(* IEC 61131-3 sources: Caravan/Archiv/12-04-19/Stations/MachineControl/MachineControl/Class/SafetyCDIAS_Base (part 6) *)

END_FUNCTION

FUNCTION VIRTUAL SafetyCDIAS_Base::GetChannelInfo
	VAR_INPUT
		pErrorMemUser 	: ^UINT;
		pErrorMem 	: ^USINT;
		ErrorDataLength 	: INT;
	END_VAR
	VAR_OUTPUT
		StateReady 	: BOOL;
	END_VAR
  VAR
  	i   : INT;
  END_VAR

  StateReady := DiagVars.UserErrorInfoReady;

  if StateReady then
    //copy error values in UserArray
    for i := 0 to ErrorDataLength-1 do

      pErrorMemUser^ := pErrorMem^;

      //set pointer to next entry
      pErrorMemUser += sizeof(UINT);
      pErrorMem += sizeof(USINT);
    end_for;
  end_if;

END_FUNCTION
